DATA_BLOCK "GDB_ManifestTest"
{ S7_Optimized_Access := 'TRUE' }
VERSION : 0.1
NON_RETAIN
VAR
    ReadLock : Bool;
END_VAR
BEGIN
END_DATA_BLOCK
